TYPE ST_EL4xx8 :
STRUCT
	ch1		:INT;
	ch2		:INT;
	ch3		:INT;
	ch4		:INT;
	ch5		:INT;
	ch6		:INT;
	ch7		:INT;
	ch8		:INT;
END_STRUCT
END_TYPE

(* stored: Version 1.1.0.1, ProductVersion 3.1.4024.12
   DUT ST_EL4xx8: Id {aadf357d-ebcd-4608-87e4-15e56b24cfb8} *)
